Fanuc KAREL source: kb00152.KL

-- PROVISIONAL review KL for V1013-1; original PC SHA256 1707429355f67cb5534d07cb1a48c51f4c48e4b3e1bf5ff4ec6834ec7e0c75d9
-- Incomplete behavior may be omitted. Consult companion uncertainty JSON. Do not deploy.
PROGRAM KB00152
%NOLOCKGROUP
VAR
  P1 : REAL
  RESULT : INTEGER
BEGIN
  -- UNRESOLVED_PC offsets 5-16; opcodes 2E,23
  -- UNRESOLVED_PC offsets 21-36; opcodes 27,22,76,23
  -- UNRESOLVED_PC offsets 41-45; opcodes 7F
END KB00152
